// TIA Portal V21 export
// export: Created 2026-10-16T07:58:28.4846108Z, ExportSetting WithDefaults, DisplayName Totally Integrated Automation Portal, DisplayVersion V21 Update 2, DisplayName TIA Portal Test Suite Advanced, DisplayVersion V21, DisplayName SINAMICS Startdrive Advanced, DisplayVersion V21 HF2, DisplayName SINAMICS DCC, DisplayVersion V21, DisplayName SINAMICS Startdrive G110M, G120, G120C, G120D, G120P, G115D, DisplayVersion V21 HF2, DisplayName SINAMICS Startdrive G130, G150, S120, S150, G200, G220, S200, S210, S220, Innomotics MVD, DisplayVersion V21 HF2, DisplayName STEP 7 Professional, DisplayVersion V21 Update 2, DisplayName STEP 7 Safety, DisplayVersion V21, DisplayName Tech WebApplication, DisplayVersion V21, DisplayName WinCC Basic/Comfort/Advanced, DisplayVersion V21 Update 2, DisplayName WinCC Unified, DisplayVersion V21 Update 2
FUNCTION_BLOCK "GraphQualification"   // FB1, GRAPH
VERSION : 0.1
// stored: AcknowledgeErrorsRequired true, AutoNumber true, GraphVersion 6.0, InitialValuesAcquisition false, IsIECCheckEnabled false, LanguageInNetworks LAD, LockOperatingMode false, PermanentILProcessingInMANMode false, SetENOAutomatically false, SkipSteps false, UDAEnableTagReadback false, WithAlarmHandling true
   // inherited from GRAPH_BASE
   VAR
      OFF_SQ_BASE : Bool;
   END_VAR
   VAR_INPUT
      ACK_EF : Bool := false;   // Alle Fehler und Störungen quittieren / Acknowledge all errors and faults
      StartCommand : Bool;
      ResetCommand : Bool;
      GuardClosed : Bool;
      SupervisionTrip : Bool;
   END_VAR
   VAR_OUTPUT
      MotorA : Bool;
      MotorB : Bool;
   END_VAR
BEGIN
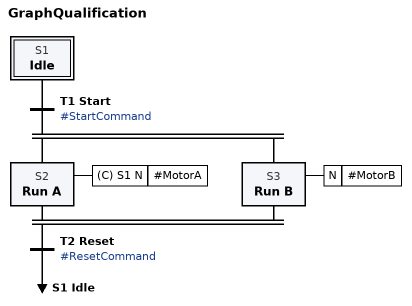
   // sequencer 1: Paralleler Ablauf / Parallel cycle
   INITIAL_STEP Idle:   // S1, max time T#10S, warning time T#7S
      interlock C := #GuardClosed;
      supervision V := #SupervisionTrip;
   END_STEP
   TRANSITION Start FROM Idle TO ("Run A", "Run B")   // T1
      := #StartCommand;
   END_TRANSITION
   STEP "Run A":   // S2, max time T#10S, warning time T#8s
      interlock C := #GuardClosed;
      supervision V := #SupervisionTrip;   // Travel timeout
      (C) S1  N    #MotorA
   END_STEP
   STEP "Run B":   // S3, max time T#10S, warning time T#7S
      interlock C := #GuardClosed;
      supervision V := #SupervisionTrip;
              N    #MotorB
   END_STEP
   TRANSITION Reset FROM ("Run A", "Run B") TO Idle   // T2, jump
      := #ResetCommand;
   END_TRANSITION
END_FUNCTION_BLOCK
